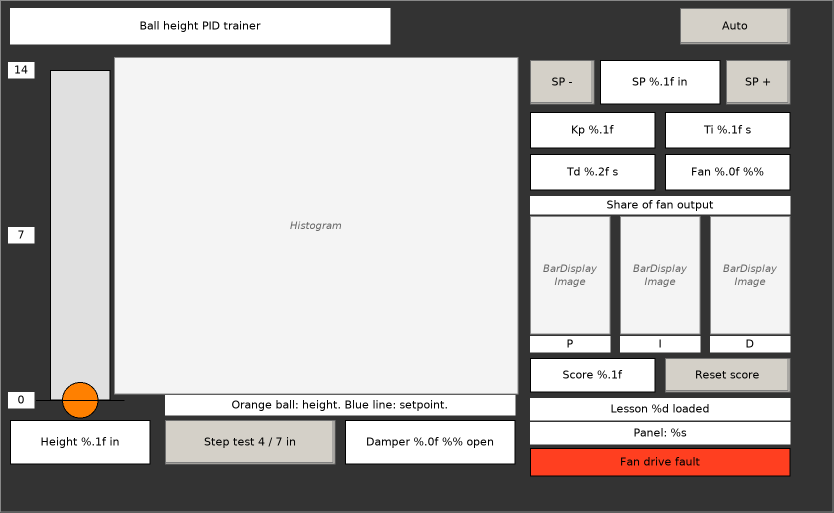
VISUALIZATION Visu_Main  // 834x513
    Rectangle (10,8 380x36), "Ball height PID trainer"
    Button (680,8 110x36), "Auto", colour toggle: P_Loop.bAuto
        toggle P_Loop.bAuto
    Rectangle (50,70 60x330)
    Ellipse (62,382 36x36)
        p2738717112: P_Hmi.nBallDY
    Line (36,400) (124,400)
        p2738717112: P_Hmi.nSPDY
    Rectangle (8,62 26x16), "14"
    Rectangle (8,227 26x16), "7"
    Rectangle (8,392 26x16), "0"
    Rectangle (10,420 140x44), "Height %.1f in", text variable: P_Hmi.rPVShow
    Rectangle (165,395 350x20), "Orange ball: height. Blue line: setpoint."
    Button (165,420 170x44), "Step test 4 / 7 in"
        tap P_Hmi.bStepTest
    Rectangle (345,420 170x44), "Damper %.0f %% open", text variable: P_Panel.rDamperPct
    Button (530,60 64x44), "SP -"
        tap P_Hmi.bSPDown
    Rectangle (600,60 120x44), "SP %.1f in", text variable: P_Loop.rSP
    Button (726,60 64x44), "SP +"
        tap P_Hmi.bSPUp
    Rectangle (530,112 125x36), "Kp %.1f", text variable: P_Loop.rKp
        OnMouseClick: write P_Loop.rKp via Default, min 0, max 20
    Rectangle (665,112 125x36), "Ti %.1f s", text variable: P_Loop.rTi
        OnMouseClick: write P_Loop.rTi via Default, min 0, max 30
    Rectangle (530,154 125x36), "Td %.2f s", text variable: P_Loop.rTd
        OnMouseClick: write P_Loop.rTd via Default, min 0, max 2
    Rectangle (665,154 125x36), "Fan %.0f %%", text variable: P_Loop.rCV
    Rectangle (530,196 260x18), "Share of fan output"
    BarDisplayImage (530,216 80x118), value: P_Hmi.rPShare, style: BarDisplayImage-Gray, scale format: %.0f, scale 0..100
    BarDisplayImage (620,216 80x118), value: P_Hmi.rIShare, style: BarDisplayImage-Gray, scale format: %.0f, scale 0..100
    BarDisplayImage (710,216 80x118), value: P_Hmi.rDShare, style: BarDisplayImage-Gray, scale format: %.0f, scale 0..100
    Rectangle (530,336 80x16), "P"
    Rectangle (620,336 80x16), "I"
    Rectangle (710,336 80x16), "D"
    Rectangle (530,358 125x34), "Score %.1f", text variable: P_Loop.rIAE
    Button (665,358 125x34), "Reset score"
        tap P_Loop.bResetIAE
    Rectangle (530,398 260x22), "Lesson %d loaded", text variable: P_Hmi.nLesson
    Rectangle (530,422 260x22), "Panel: %s", text variable: P_Panel.sState
    Rectangle (530,448 260x28), "Fan drive fault", invisible if: NOT P_Panel.bFanFault
    Histogram (114,57 404x337), scale format: %.0f, scale 0..14
        p1518820177: P_Hmi.aTrendPV
        p102497268: P_Hmi.aTrendPV
        p788070771: ARRAY [0..149] OF REAL
    Potentiometer360 (834,512 0x1), style: Potentiometer-Potentiometer360-Gray, scale format: %.1f, scale 0..100
        p2431819421: Outside
END_VISUALIZATION

(* stored: Version 1.1.0.1
   Visu Visu_Main: Id {c6a46cf5-3522-40de-972d-9aa613973555} *)
